(* IEC 61131-3 sources: guidance-for-physical-ai-production-designer-on-aws/source/plan2cell/examples/welding_cell_2_small/plc/trust/head/src (part 2) *)

(* ---- FB_ZoneArbiter.st ---- *)
(*
 * FB_ZoneArbiter
 * Generated by bt2plc 0.1.0 for cell welding_cell_2_small (plan bt_1790934549_welding_cell_2_small)
 *
 * Zone (mutex) and permit arbiter, data-driven by GVL_Cell (aTickets, anZoneFirst/Count,
 * aOps[].dwZoneMask / nPredFirst / nPredCount, aPreds).
 *
 * REQUEST / GRANT DWORD: bits 0..30 = zones 1..31, bit 31 = PERMIT (GVL_Cell.PERMIT_MASK).
 *   GP_PLANNED : a zone is granted only to its next ticket holder, only if the request
 *                equals the op's full mask and the reported op index matches the ticket.
 *   GP_FCFS    : free zones to any requester whose request equals the op mask, oldest
 *                request first, ties by robot index; zones of an older requester that
 *                waits only for occupied zones are reserved against younger ones.
 *                BT ordering is NOT preserved by the zones.
 *   PERMIT     : granted for op (r, k) iff every pred (q, j) of the op has anDone[q] >= j.
 *                Not a mutex: never held against other robots, released when bit 31 drops.
 * Both policies grant all bits of an op in the same scan (all-or-nothing).
 *
 * Checks: 4-phase handshake (op index must not change while a grant is held), release
 * only by a robot that runs OK, holder raising extra bits; request mask and ticket checks
 * are evaluated once (op index, REQUEST) has been stable for tDebounce.
 * Fail closed: any violation latches bFault and drops all grants until bReset.
 *
 * Timing uses tNow (monotonic TIME from the caller's clock), no timer instances.
 *)

FUNCTION_BLOCK FB_ZoneArbiter
VAR_INPUT
    bReset              : BOOL;             (* Level: rewind tickets, clear holders, grants and fault *)
    bEnable             : BOOL;             (* New grants allowed *)
    ePolicy             : E_GrantPolicy := E_GrantPolicy#GP_PLANNED;
    tDebounce           : TIME := T#200MS;  (* (op index, REQUEST) stable time before mask / ticket checks *)
    tNow                : TIME;             (* Monotonic time of this scan *)
    abRobotOk           : ARRAY[1..2] OF BOOL;      (* Production job running, no robot error *)
    awStep              : ARRAY[1..2] OF WORD;      (* Reported op index, 0 = none *)
    adwReq              : ARRAY[1..2] OF DWORD;     (* REQUEST DWORD *)
    anDone              : ARRAY[1..2] OF INT;       (* Ops completed per robot in this cycle *)
END_VAR

VAR_OUTPUT
    adwGrant            : ARRAY[1..2] OF DWORD;     (* GRANT DWORD per robot *)
    anHolder            : ARRAY[1..2] OF INT;    (* Robot holding the zone, 0 = free *)
    anTicket            : ARRAY[1..2] OF INT;    (* Next ticket index in GVL_Cell.aTickets *)
    bAllConsumed        : BOOL;             (* No zone held and (planned) every ticket consumed *)
    bFault              : BOOL;
    eFault              : E_CellError;
    nFaultRobot         : INT;
    nFaultZone          : INT;
END_VAR

VAR
    _udiScan            : UDINT;            (* Scan counter: request age for FCFS *)
    _audiWaitSince      : ARRAY[1..2] OF UDINT;     (* Scan of the first pending request, 0 = none *)
    _abPicked           : ARRAY[1..2] OF BOOL;
    _anGrantStep        : ARRAY[1..2] OF INT;       (* Op index at the time of the grant *)
    _awPrevStep         : ARRAY[1..2] OF WORD;
    _adwPrevReq         : ARRAY[1..2] OF DWORD;
    _atChange           : ARRAY[1..2] OF TIME;      (* tNow of the last (op index, REQUEST) change *)
    _abStable           : ARRAY[1..2] OF BOOL;
    _eNew               : E_CellError;
    _nNewRobot          : INT;
    _nNewZone           : INT;
    _k                  : INT;
    _r                  : INT;
    _rr                 : INT;
    _rSel               : INT;
    _z                  : INT;
    _p                  : INT;
    _q                  : INT;
    _iOp                : INT;
    _nStep              : INT;
    _nTicket            : INT;
    _nLastTicket        : INT;
    _nPredFirst         : INT;
    _nPredLast          : INT;
    _dwBit              : DWORD;
    _dwExp              : DWORD;            (* Expected REQUEST of the reported op *)
    _dwZones            : DWORD;            (* Zone bits of _dwExp (permit bit removed) *)
    _dwReserved         : DWORD;            (* FCFS: zones reserved by older requesters this scan *)
    _bOk                : BOOL;             (* All zones of the op grantable *)
    _bPermitOk          : BOOL;             (* All permit predecessors done *)
    _bPending           : BOOL;
END_VAR
(*
 * FB_ZoneArbiter - Implementation
 * Order per scan: debounce + handshake check, release, grant, fault latch.
 *)

IF bReset THEN
    FOR _z := 1 TO GVL_Cell.N_ZONES DO
        anHolder[_z] := 0;
        anTicket[_z] := GVL_Cell.anZoneFirst[_z];
    END_FOR
    FOR _r := 1 TO GVL_Cell.N_ROBOTS DO
        adwGrant[_r] := DWORD#0;
        _audiWaitSince[_r] := 0;
        _anGrantStep[_r] := 0;
        _awPrevStep[_r] := awStep[_r];
        _adwPrevReq[_r] := adwReq[_r];
        _atChange[_r] := tNow;
        _abStable[_r] := FALSE;
    END_FOR
    _udiScan := 0;
    bFault := FALSE;
    eFault := E_CellError#ERR_NONE;
    nFaultRobot := 0;
    nFaultZone := 0;
    bAllConsumed := (GVL_Cell.N_ZONES = 0) OR (ePolicy = E_GrantPolicy#GP_FCFS);
    RETURN;
END_IF

IF bFault THEN
    RETURN;                                 (* latched until bReset *)
END_IF

_udiScan := _udiScan + 1;
_eNew := E_CellError#ERR_NONE;
_nNewRobot := 0;
_nNewZone := 0;

(* ============================================================================
   0. DEBOUNCE / 4-PHASE HANDSHAKE
   ============================================================================ *)
FOR _r := 1 TO GVL_Cell.N_ROBOTS DO
    IF (awStep[_r] <> _awPrevStep[_r]) OR (adwReq[_r] <> _adwPrevReq[_r]) THEN
        _atChange[_r] := tNow;
        _awPrevStep[_r] := awStep[_r];
        _adwPrevReq[_r] := adwReq[_r];
    END_IF
    _abStable[_r] := (tNow - _atChange[_r]) >= tDebounce;

    (* A correct robot changes its op index only after it has seen GRANT = 0. Profile vw-ks24
       has no 4-phase handshake: there the robot only holds its release level long enough for
       the head to see it (bt2krl emits a dwell after every release), so the check needs the
       debounce to avoid firing on scan jitter. *)
    IF (adwGrant[_r] <> DWORD#0) AND (WORD_TO_INT(awStep[_r]) <> _anGrantStep[_r])
       AND (_abStable[_r] OR NOT GVL_Cell.PROFILE_VW)
       AND (_eNew = E_CellError#ERR_NONE) THEN
        _eNew := E_CellError#ERR_HANDSHAKE;
        _nNewRobot := _r;
        _nNewZone := 0;
    END_IF
END_FOR

(* ============================================================================
   1. RELEASE - holder dropped its REQUEST bit
   ============================================================================ *)
FOR _z := 1 TO GVL_Cell.N_ZONES DO
    _rr := anHolder[_z];
    IF _rr <> 0 THEN
        _dwBit := SHL(DWORD#1, _z - 1);
        IF (adwReq[_rr] AND _dwBit) = DWORD#0 THEN
            IF abRobotOk[_rr] THEN
                anHolder[_z] := 0;
                adwGrant[_rr] := adwGrant[_rr] AND NOT _dwBit;
                IF ePolicy = E_GrantPolicy#GP_PLANNED THEN
                    anTicket[_z] := anTicket[_z] + 1;
                END_IF
            ELSIF _eNew = E_CellError#ERR_NONE THEN
                (* request vanished because the robot stopped / faulted / lost
                   connection: the zone may still be occupied - never re-grant *)
                _eNew := E_CellError#ERR_RELEASE_INVALID;
                _nNewRobot := _rr;
                _nNewZone := _z;
            END_IF
        END_IF
    END_IF
END_FOR

(* Permit bit: not a mutex, released as soon as REQUEST bit 31 drops *)
FOR _r := 1 TO GVL_Cell.N_ROBOTS DO
    IF ((adwGrant[_r] AND GVL_Cell.PERMIT_MASK) <> DWORD#0)
       AND ((adwReq[_r] AND GVL_Cell.PERMIT_MASK) = DWORD#0) THEN
        adwGrant[_r] := adwGrant[_r] AND NOT GVL_Cell.PERMIT_MASK;
    END_IF
END_FOR

(* ============================================================================
   2. GRANT
   ============================================================================ *)
FOR _r := 1 TO GVL_Cell.N_ROBOTS DO
    _abPicked[_r] := FALSE;
    IF (adwReq[_r] = DWORD#0) OR (adwGrant[_r] <> DWORD#0) THEN
        _audiWaitSince[_r] := 0;
    ELSIF _audiWaitSince[_r] = 0 THEN
        _audiWaitSince[_r] := _udiScan;
    END_IF
END_FOR
_dwReserved := DWORD#0;

FOR _k := 1 TO GVL_Cell.N_ROBOTS DO
    (* --- visiting order: PLANNED = robot index, FCFS = oldest request first --- *)
    _rSel := 0;
    FOR _r := 1 TO GVL_Cell.N_ROBOTS DO
        IF NOT _abPicked[_r] THEN
            IF _rSel = 0 THEN
                _rSel := _r;
            ELSIF (ePolicy = E_GrantPolicy#GP_FCFS) AND (_audiWaitSince[_r] <> 0) THEN
                IF (_audiWaitSince[_rSel] = 0) OR (_audiWaitSince[_r] < _audiWaitSince[_rSel]) THEN
                    _rSel := _r;
                END_IF
            END_IF
        END_IF
    END_FOR
    _rr := _rSel;
    _abPicked[_rr] := TRUE;

    (* --- expected mask of the op the robot reports --- *)
    _nStep := WORD_TO_INT(awStep[_rr]);
    _iOp := 0;
    _dwExp := DWORD#0;
    IF (_nStep >= 1) AND (_nStep <= GVL_Cell.anRobotOpCount[_rr]) THEN
        _iOp := GVL_Cell.anRobotFirstOp[_rr] + _nStep - 1;
        _dwExp := GVL_Cell.aOps[_iOp].dwZoneMask;
    END_IF
    _dwZones := _dwExp AND NOT GVL_Cell.PERMIT_MASK;

    _bPending := bEnable AND abRobotOk[_rr] AND (adwReq[_rr] <> DWORD#0) AND (adwGrant[_rr] = DWORD#0);

    (* --- request must equal the op mask (debounced) --- *)
    IF _bPending AND _abStable[_rr] AND (adwReq[_rr] <> _dwExp)
       AND (_eNew = E_CellError#ERR_NONE) THEN
        _eNew := E_CellError#ERR_REQ_MISMATCH;
        _nNewRobot := _rr;
        _nNewZone := 0;
    END_IF

    (* --- a holder must not raise bits it was not granted --- *)
    IF (adwGrant[_rr] <> DWORD#0) AND ((adwReq[_rr] AND NOT adwGrant[_rr]) <> DWORD#0)
       AND (_eNew = E_CellError#ERR_NONE) THEN
        _eNew := E_CellError#ERR_UNEXPECTED_REQUEST;
        _nNewRobot := _rr;
        _nNewZone := 0;
    END_IF

    IF _bPending AND (adwReq[_rr] = _dwExp) THEN
        (* --- zones: all free, (planned) ticket = this op, (FCFS) not reserved --- *)
        _bOk := TRUE;
        FOR _z := 1 TO GVL_Cell.N_ZONES DO
            _dwBit := SHL(DWORD#1, _z - 1);
            IF (_dwZones AND _dwBit) <> DWORD#0 THEN
                IF anHolder[_z] <> 0 THEN
                    _bOk := FALSE;
                ELSIF ePolicy = E_GrantPolicy#GP_PLANNED THEN
                    _nTicket := anTicket[_z];
                    _nLastTicket := GVL_Cell.anZoneFirst[_z] + GVL_Cell.anZoneCount[_z] - 1;
                    IF (_nTicket < GVL_Cell.anZoneFirst[_z]) OR (_nTicket > _nLastTicket) THEN
                        _bOk := FALSE;              (* zone consumed *)
                        IF _abStable[_rr] AND (_eNew = E_CellError#ERR_NONE) THEN
                            _eNew := E_CellError#ERR_TICKET_SKIPPED;
                            _nNewRobot := _rr;
                            _nNewZone := _z;
                        END_IF
                    ELSIF (GVL_Cell.aTickets[_nTicket].nRobot <> _rr)
                          OR (GVL_Cell.aTickets[_nTicket].nOp <> _nStep) THEN
                        _bOk := FALSE;              (* not this op's turn yet *)
                        IF (GVL_Cell.aTickets[_nTicket].nRobot = _rr) AND _abStable[_rr]
                           AND (_eNew = E_CellError#ERR_NONE) THEN
                            _eNew := E_CellError#ERR_TICKET_SKIPPED;
                            _nNewRobot := _rr;
                            _nNewZone := _z;
                        END_IF
                    END_IF
                ELSIF (_dwReserved AND _dwBit) <> DWORD#0 THEN
                    _bOk := FALSE;                  (* FCFS: reserved by an older requester *)
                END_IF
            END_IF
        END_FOR

        (* --- permit: every predecessor op done --- *)
        _bPermitOk := TRUE;
        IF ((_dwExp AND GVL_Cell.PERMIT_MASK) <> DWORD#0) AND (_iOp >= 1) THEN
            (* GVL array elements are copied to locals before use as call arguments *)
            _nPredFirst := GVL_Cell.aOps[_iOp].nPredFirst;
            _nPredLast := _nPredFirst + GVL_Cell.aOps[_iOp].nPredCount - 1;
            _nPredFirst := MAX(1, _nPredFirst);
            _nPredLast := MIN(GVL_Cell.N_PREDS, _nPredLast);
            FOR _p := _nPredFirst TO _nPredLast DO
                _q := GVL_Cell.aPreds[_p].nRobot;
                IF (_q < 1) OR (_q > GVL_Cell.N_ROBOTS) THEN
                    _bPermitOk := FALSE;
                ELSIF anDone[_q] < GVL_Cell.aPreds[_p].nOp THEN
                    _bPermitOk := FALSE;
                END_IF
            END_FOR
        END_IF

        IF _bOk AND _bPermitOk THEN
            FOR _z := 1 TO GVL_Cell.N_ZONES DO
                IF (_dwZones AND SHL(DWORD#1, _z - 1)) <> DWORD#0 THEN
                    anHolder[_z] := _rr;
                END_IF
            END_FOR
            adwGrant[_rr] := _dwExp;
            _anGrantStep[_rr] := _nStep;
            _audiWaitSince[_rr] := 0;
        ELSIF _bPermitOk AND (ePolicy = E_GrantPolicy#GP_FCFS) THEN
            (* older requester blocked only by occupied / reserved zones: reserve them
               (a requester still waiting for its permit reserves nothing - no deadlock) *)
            _dwReserved := _dwReserved OR _dwZones;
        END_IF
    END_IF
END_FOR

(* ============================================================================
   3. FAULT LATCH / CYCLE COMPLETENESS
   ============================================================================ *)
IF _eNew <> E_CellError#ERR_NONE THEN
    bFault := TRUE;
    eFault := _eNew;
    nFaultRobot := _nNewRobot;
    nFaultZone := _nNewZone;
    FOR _r := 1 TO GVL_Cell.N_ROBOTS DO
        adwGrant[_r] := DWORD#0;
    END_FOR
END_IF

bAllConsumed := TRUE;
FOR _z := 1 TO GVL_Cell.N_ZONES DO
    IF anHolder[_z] <> 0 THEN
        bAllConsumed := FALSE;
    ELSIF (ePolicy = E_GrantPolicy#GP_PLANNED)
          AND (anTicket[_z] <= GVL_Cell.anZoneFirst[_z] + GVL_Cell.anZoneCount[_z] - 1) THEN
        bAllConsumed := FALSE;
    END_IF
END_FOR
END_FUNCTION_BLOCK

(* ---- PLC_PRG.st ---- *)
(*
 * PLC_PRG - Head PLC cell program
 * Generated by bt2plc 0.1.0 for cell welding_cell_2_small (plan bt_1790934549_welding_cell_2_small)
 *
 * Copies every robot's GVL_IO block into the cell's input array, runs FB_Cell and
 * copies the commands back (whole arrays / single bytes only).
 *
 * Operator (plain VARs, pulses are cleared after each scan):
 *   bAutoRun          Level: start a cycle whenever the cell is READY
 *                     (initialised from GVL_Cell.AUTO_RUN on the first scan)
 *   bStart            Pulse: start one cycle
 *   bStop             Pulse: abort (ERR_OPERATOR_STOP); latched in every state, also
 *                     cancels a running reset (CS_RESETTING -> CS_ERROR)
 *   bReset            Pulse: reset after an error (a pulse during CS_ABORTING is kept)
 *   bRecoveryConfirm  Pulse: after an abort mid-cycle or a start-up with an active robot
 *                     away from home, robots moved clear -> sequential blind homing
 *
 * Status: PLC_PRG.fbCell.eState / eError / nErrorRobot / nErrorOp / nErrorZone /
 *         bRecoveryRequired / udiCycles / tLastCycle / aeRobotState / awStep / adwGrant ...
 *
 * Task: MainTask (4 ms cycle)
 *)

PROGRAM PLC_PRG
VAR
    (* Cell controller *)
    fbCell              : FB_Cell;

    (* === Operator === *)
    bAutoRun            : BOOL := TRUE;     (* overwritten by GVL_Cell.AUTO_RUN on the first scan *)
    bStart              : BOOL;
    bStop               : BOOL;
    bReset              : BOOL;
    bRecoveryConfirm    : BOOL;

    (* === Status readback === *)
    eCellState          : E_CellState;
    eCellError          : E_CellError;
    bCellError          : BOOL;
    bRecoveryRequired   : BOOL;
    udiCycles           : UDINT;

    (* Robot input images for fbCell *)
    _astIn              : ARRAY[1..2] OF ST_RobotIn;
    _bFirstScan         : BOOL := TRUE;
END_VAR
(*
 * PLC_PRG - Implementation
 *)

IF _bFirstScan THEN
    bAutoRun := GVL_Cell.AUTO_RUN;
    _bFirstScan := FALSE;
END_IF

(* ============================================================================
   INPUTS: GVL_IO -> fbCell (robot -> PLC)
   ============================================================================ *)

(* 1: R1 - robot1 - kuka_robi1 (kuka-robi1, 192.168.100.11) *)
_astIn[1].abySafeIn[0] := GVL_IO.bySafeIn0_R1;
_astIn[1].abySafeIn[1] := GVL_IO.bySafeIn1_R1;
_astIn[1].abySafeIn[2] := GVL_IO.bySafeIn2_R1;
_astIn[1].abySafeIn[3] := GVL_IO.bySafeIn3_R1;
_astIn[1].abySafeIn[4] := GVL_IO.bySafeIn4_R1;
_astIn[1].abySafeIn[5] := GVL_IO.bySafeIn5_R1;
_astIn[1].abySafeIn[6] := GVL_IO.bySafeIn6_R1;
_astIn[1].abySafeIn[7] := GVL_IO.bySafeIn7_R1;
_astIn[1].aVassIn := GVL_IO.aVassInputData_R1;

(* 2: R2 - robot2 - kuka_robi2 (kuka-robi2, 192.168.100.12) *)
_astIn[2].abySafeIn[0] := GVL_IO.bySafeIn0_R2;
_astIn[2].abySafeIn[1] := GVL_IO.bySafeIn1_R2;
_astIn[2].abySafeIn[2] := GVL_IO.bySafeIn2_R2;
_astIn[2].abySafeIn[3] := GVL_IO.bySafeIn3_R2;
_astIn[2].abySafeIn[4] := GVL_IO.bySafeIn4_R2;
_astIn[2].abySafeIn[5] := GVL_IO.bySafeIn5_R2;
_astIn[2].abySafeIn[6] := GVL_IO.bySafeIn6_R2;
_astIn[2].abySafeIn[7] := GVL_IO.bySafeIn7_R2;
_astIn[2].aVassIn := GVL_IO.aVassInputData_R2;

(* ============================================================================
   CELL
   ============================================================================ *)
fbCell(
    bEnable             := TRUE,
    bAutoRun            := bAutoRun,
    bStart              := bStart,
    bStop               := bStop,
    bReset              := bReset,
    bRecoveryConfirm    := bRecoveryConfirm,
    astIn               := _astIn,
    eState              => eCellState,
    eError              => eCellError,
    bError              => bCellError,
    bRecoveryRequired   => bRecoveryRequired,
    udiCycles           => udiCycles);

(* ============================================================================
   OUTPUTS: fbCell -> GVL_IO (PLC -> robot)
   ============================================================================ *)

(* 1: R1 - robot1 *)
GVL_IO.bySafeOut0_R1 := fbCell.astOut[1].abySafeOut[0];
GVL_IO.bySafeOut1_R1 := fbCell.astOut[1].abySafeOut[1];
GVL_IO.bySafeOut2_R1 := fbCell.astOut[1].abySafeOut[2];
GVL_IO.bySafeOut3_R1 := fbCell.astOut[1].abySafeOut[3];
GVL_IO.bySafeOut4_R1 := fbCell.astOut[1].abySafeOut[4];
GVL_IO.bySafeOut5_R1 := fbCell.astOut[1].abySafeOut[5];
GVL_IO.bySafeOut6_R1 := fbCell.astOut[1].abySafeOut[6];
GVL_IO.bySafeOut7_R1 := fbCell.astOut[1].abySafeOut[7];
GVL_IO.aVassOutputData_R1 := fbCell.astOut[1].aVassOut;

(* 2: R2 - robot2 *)
GVL_IO.bySafeOut0_R2 := fbCell.astOut[2].abySafeOut[0];
GVL_IO.bySafeOut1_R2 := fbCell.astOut[2].abySafeOut[1];
GVL_IO.bySafeOut2_R2 := fbCell.astOut[2].abySafeOut[2];
GVL_IO.bySafeOut3_R2 := fbCell.astOut[2].abySafeOut[3];
GVL_IO.bySafeOut4_R2 := fbCell.astOut[2].abySafeOut[4];
GVL_IO.bySafeOut5_R2 := fbCell.astOut[2].abySafeOut[5];
GVL_IO.bySafeOut6_R2 := fbCell.astOut[2].abySafeOut[6];
GVL_IO.bySafeOut7_R2 := fbCell.astOut[2].abySafeOut[7];
GVL_IO.aVassOutputData_R2 := fbCell.astOut[2].aVassOut;

(* One-shot operator buttons *)
bStart := FALSE;
bStop := FALSE;
bReset := FALSE;
bRecoveryConfirm := FALSE;
END_PROGRAM
